{region 'Documentation'}
(*!
<summary>Check equality between consecutive active observations.</summary>
<description>

The first active observation establishes a baseline without deciding a result. Disabling
observation invalidates that baseline, not the held Result. Re-enabling first establishes a new
baseline; Reset clears history.

ObserveFirstCycle FALSE delays the first observation by one enabled call.

</description>
*)
{endregion}
FUNCTION_BLOCK AssertNoValueChange_USInt EXTENDS AssertionBase
VAR_INPUT
    IN : USINT; //! Actual value to observe.
END_VAR
VAR
    FINPrevious : USINT;
    FObservationPrevious : BOOL;
    FEvaluationActive : BOOL;
END_VAR

SUPER^();

{region 'Documentation'}
(*!
<summary>Observe the current value before evaluating a change against the previous observation.</summary>
*)
{endregion}
METHOD PROTECTED Assert
VAR
    PreviousValue : USINT;
    Message : STRING(GVL_Constants.MessageLength);
    PreviousText : STRING(GVL_Constants.AssertionValueLength);
    ActualText : STRING(GVL_Constants.AssertionValueLength);
END_VAR
FEvaluationActive := ObservationActive AND FObservationPrevious;
FObservationPrevious := ObservationActive;

IF NOT ObservationActive THEN
    RETURN;
END_IF;

PreviousValue := FINPrevious;
FINPrevious := IN;

IF NOT EvaluationActive THEN
    RETURN;
END_IF;

IF Result = E_Result.Error THEN
    RETURN;
END_IF;

IF Result = E_Result.Failed THEN
    RETURN;
END_IF;

IF IN <> PreviousValue THEN
    PreviousText := USINT_TO_STRING(PreviousValue);
    ActualText := USINT_TO_STRING(IN);
    Message := CONCAT('Assertion failed: value changed unexpectedly. Previous = ',
        PreviousText);
    Message := CONCAT(Message, ', Actual = ');
    Message := CONCAT(Message, ActualText);
    Message := CONCAT(Message, '.');
    Fail(Message := Message);
    RETURN;
END_IF;

Pass();
END_METHOD

{region 'Documentation'}
(*!
<summary>Current/last call has an active observation and a preceding observation
baseline.</summary>
*)
{endregion}
{attribute 'monitoring' := 'call'}
PROPERTY PUBLIC EvaluationActive : BOOL //! Current/last call has an active observation and a preceding observation baseline.
GET // PUBLIC
EvaluationActive := FEvaluationActive;
END_GET
END_PROPERTY

{region 'Documentation'}
(*!
<summary>Clear observation history and the current evaluation gate.</summary>
*)
{endregion}
METHOD PROTECTED ResetAssertion
FINPrevious := 0;
FObservationPrevious := FALSE;
FEvaluationActive := FALSE;
END_METHOD

END_FUNCTION_BLOCK

(* stored: Version 1.1.0.1
   POU AssertNoValueChange_USInt: Id {a48bf548-85b0-40f4-ab25-c64f1e64616b}, SpecialFunc None
   Folder Internal: Id {36861742-a85e-4cbc-a7a5-ed38e0992c3e}
   Method Assert: Id {31f28491-44ca-42e4-98d9-efd0ad607406}
   Property EvaluationActive: Id {92f170f9-271a-4a63-be9d-00bb7ca193bc}
   Get Get: Id {5be0bc11-c9b4-4834-85e0-3deb9afa87f7}
   Method ResetAssertion: Id {a699a017-1110-4844-adf3-fb9a9d7adcb5} *)
